Yaskawa INFORM job: TGTPROG.JBI

/JOB
//NAME TGTPROG
//POS
///NPOS 3,0,0,0,0,0
///TOOL 9
///POSTYPE PULSE
///PULSE
C00000=10,-20,30,-40,50,-60
C00001=0,0,0,2,-3,3
C00002=0,1,-2,2,0,0
//INST
<volatile>
///COMM Generated using RoboDK
///ATTR SC,RW
///GROUP1 RB1
NOP
'Program generated by RoboDK v
'6.0.7 for Yaskawa Motoman GP8
' on XX/XX/XXXX 18:00:00
'Using nominal kinematics.
MOVJ C00000 VJ=50.00
MOVL C00001 V=100.0
MOVJ C00002 VJ=50.00
END
